TYPE "DT_REFERENCE_ALL"
VERSION : 0.1
   STRUCT
      WATER_LEVEL : "DT_REFERENCE_SOLO";
      GATE_1 : "DT_REFERENCE_SOLO";
      GATE_2 : "DT_REFERENCE_SOLO";
      GATE_3 : "DT_REFERENCE_SOLO";
      GATE_4 : "DT_REFERENCE_SOLO";
      GATE_5 : "DT_REFERENCE_SOLO";
      GATE_6 : "DT_REFERENCE_SOLO";
      GATE_7 : "DT_REFERENCE_SOLO";
      GATE_8 : "DT_REFERENCE_SOLO";
      GATE_9 : "DT_REFERENCE_SOLO";
      GATE_10 : "DT_REFERENCE_SOLO";
      SPARE_11 : "DT_REFERENCE_SOLO";
      SPARE_12 : "DT_REFERENCE_SOLO";
      SPARE_13 : "DT_REFERENCE_SOLO";
      SPARE_14 : "DT_REFERENCE_SOLO";
      SPARE_15 : "DT_REFERENCE_SOLO";
      SPARE_16 : "DT_REFERENCE_SOLO";
      SPARE_17 : "DT_REFERENCE_SOLO";
      SPARE_18 : "DT_REFERENCE_SOLO";
      SPARE_19 : "DT_REFERENCE_SOLO";
      SPARE_20 : "DT_REFERENCE_SOLO";
      SPARE_21 : "DT_REFERENCE_SOLO";
      SPARE_22 : "DT_REFERENCE_SOLO";
      SPARE_23 : "DT_REFERENCE_SOLO";
      SPARE_24 : "DT_REFERENCE_SOLO";
      SPARE_25 : "DT_REFERENCE_SOLO";
      SPARE_26 : "DT_REFERENCE_SOLO";
      SPARE_27 : "DT_REFERENCE_SOLO";
      SPARE_28 : "DT_REFERENCE_SOLO";
      SPARE_29 : "DT_REFERENCE_SOLO";
      SPARE_30 : "DT_REFERENCE_SOLO";
      SPARE_31 : "DT_REFERENCE_SOLO";
   END_STRUCT;

END_TYPE

